Yaskawa INFORM job: SPLITTE.JBI

/JOB
//NAME SPLITTE
//POS
///NPOS 5,0,0,0,0,0
///TOOL 1
///POSTYPE PULSE
///PULSE
C00000=10,20,-10,30,-45,60
C00001=18,24,-10,30,-45,60
C00002=14,20,-5,30,-45,60
C00003=18,24,-10,30,-45,60
C00004=14,20,-5,30,-45,60
//INST
///DATE 2026/10/26 01:19
///COMM Generated using RoboDK
///ATTR SC,RW
///GROUP1 RB1
NOP
'Program generated by Vertical
'Bot Studio for Motoman GP8 on
' 25/10/2026 12:00:00
'Using nominal kinematics.
'Using Frame 2 (targets wrt ba
'se):
'100.0,-50.0,20.0,0.0,0.0,30.0
'Tool 1 (Tool 1) should be clo
'se to:
'10.0,0.0,120.0,0.0,15.0,0.0
MOVJ C00000 VJ=50.00
MOVL C00001 V=200.0
MOVL C00002 V=200.0
MOVL C00003 V=200.0
MOVL C00004 V=200.0
END
